SUBAPPLICATION AUI_GT_0 (* Prüft ob UINT-Adapter Wert > 0 ist (AX-Adapter Ausgang) *)
  (* Standard: 61499-2 *)
  (* Version 1.0, 2026-04-20, franz, Meisterschulen am Ostbahnhof *)
  PACKAGE MyLib::sys;
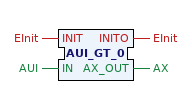
  EVENT_INPUT
    INIT : EInit; (* Initialization Request *)
  END_EVENT
  EVENT_OUTPUT
    INITO : EInit; (* Initialization Confirm *)
  END_EVENT
  SOCKETS
    IN : adapter::types::unidirectional::AUI;
  END_SOCKETS
  PLUGS
    AX_OUT : adapter::types::unidirectional::AX;
  END_PLUGS
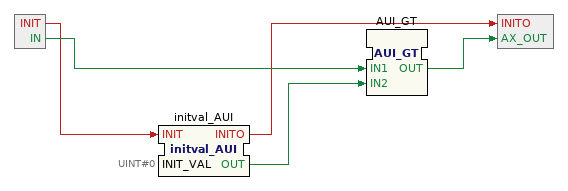
  FBS
    AUI_GT : adapter::iec61131::comparison::AUI_GT;
    initval_AUI : adapter::types::unidirectional::AUI::initval::initval_AUI(INIT_VAL := UINT#0);
  END_FBS
  EVENT_CONNECTIONS
    INIT TO initval_AUI.INIT;
    initval_AUI.INITO TO INITO;
  END_CONNECTIONS
  ADAPTER_CONNECTIONS
    IN TO AUI_GT.IN1;
    AUI_GT.OUT TO AX_OUT;
    initval_AUI.OUT TO AUI_GT.IN2;
  END_CONNECTIONS
END_SUBAPPLICATION
